// TIA Portal V21 export
// export: Created 2026-11-21T13:54:30.6197884Z, ExportSetting WithDefaults, DisplayName Totally Integrated Automation Portal, DisplayVersion V21, DisplayName STEP 7 Professional, DisplayVersion V21, DisplayName STEP 7 Safety, DisplayVersion V21, DisplayName Tech WebApplication, DisplayVersion V21, DisplayName WinCC Basic/Comfort/Advanced, DisplayVersion V21, DisplayName WinCC Unified, DisplayVersion V21
VAR_GLOBAL   // PLC tag table "Tank"
   Tank_Level AT %IW64 : Int;   // Level of the tank in percent
   Tank_Temp AT %MD20 : Real;   // Temperature of the tank
   Agitator_On AT %Q0.0 : Bool;   // The agitator runs
   Alarm_Word AT %MW30 : Word;   // Alarm bits of the mixer
END_VAR
